(*
SPDX-FileCopyrightText: © 2026 Oleksandr Tiutyk <trofimich@gmail.com>
SPDX-License-Identifier: MIT
License: https://opensource.org/license/mit
*)

(*!
<summary>
Beckhoff EL3204: 4-channel RTD resistance thermometer terminal (Pt100, Pt1000, Ni120...).
</summary>
<description>
Process image mapping structure for the EL3204 4-channel RTD temperature input terminal.
When used for I/O, link located fields or their containing buffers to the matching selected PDOs.
The record is not a packed wire buffer; compiler padding is not part of the device specification.
Unlinked/default values do not prove valid I/O. The caller evaluates bus/channel validity before use.
Use one owner task per instance and externally synchronize other access; multi-field snapshots are not atomic.
Copies store data without creating hardware links. Keep borrowed field references valid while consumers are bound.
This passive record performs no validation, synchronization, configuration or protocol advancement.
Select standard status-plus-INT16 PDOs; compact layouts are unsupported. Configure presentation explicitly:
0.1/0.01 deg C per digit follows the device setting, not this record.
</description>
*)
TYPE EL3204 :
STRUCT
	Ch1 : RTD_INPUT_CHANNEL;
	Ch2 : RTD_INPUT_CHANNEL;
	Ch3 : RTD_INPUT_CHANNEL;
	Ch4 : RTD_INPUT_CHANNEL;
END_STRUCT
END_TYPE

(* stored: Version 1.1.0.1, ProductVersion 3.1.4026.20
   DUT EL3204: Id {a8da5a93-77c5-431a-8666-6edf8676f5f7} *)
